(* IEC 61131-3 sources: Codesys_IAP/Demo/PLC1/Magazijn Overzetter Simulatie Structured Text 2V1_tekst/Programma Structured Text/StationClass, 8 files *)

(* ---- cycle.st ---- *)
(*#### DECLARATIE ####*)
// Datum : 26 november 2026, Auteur: Gerard Harkema
METHOD cycle
VAR
END_VAR
(*#### IMPLEMENTATIE ####*)
// Eerst de objecten
magazijn.cycle();
overzetter.cycle();

// Dan de fouten: een fout in een object zet het hele station in error
IF magazijn.isError() OR overzetter.isError() THEN
	eState := stationStates.error;
END_IF

// Dan de coordinatie, volgens het statediagram van StationClass
CASE eState OF
	stationStates.idle:
		; // wacht op start()

	stationStates.magazijn_uitstoten:
		IF magazijn.start() THEN		// TRUE = mislukt
			eState := stationStates.error;
		ELSE
			eState := stationStates.wacht_magazijn_klaar;
		END_IF

	stationStates.wacht_magazijn_klaar:
		IF magazijn.isKlaar() THEN
			eState := stationStates.overzetten;
		END_IF

	stationStates.overzetten:
		IF overzetter.start() THEN		// TRUE = mislukt
			eState := stationStates.error;
		ELSE
			eState := stationStates.wacht_overzetter_klaar;
		END_IF

	stationStates.wacht_overzetter_klaar:
		IF overzetter.isKlaar() THEN
			eState := stationStates.idle;
		END_IF

	stationStates.error:
		; // wacht op reset()
END_CASE

(* ---- initialize.st ---- *)
(*#### DECLARATIE ####*)
// Datum : 26 november 2026, Auteur: Gerard Harkema
METHOD initialize
VAR_INPUT
	IORef			: REFERENCE TO stationIO;
END_VAR
(*#### IMPLEMENTATIE ####*)
IO REF= IORef;

// Elk object krijgt zijn eigen IO-structuur
magazijn.initialize(IO.magazijn);
overzetter.initialize(IO.overzetter);

eState := stationStates.idle;

(* ---- isError.st ---- *)
(*#### DECLARATIE ####*)
// Datum : 26 november 2026, Auteur: Gerard Harkema
METHOD isError : BOOL
VAR_INPUT
END_VAR
(*#### IMPLEMENTATIE ####*)
isError := (eState = stationStates.error);

(* ---- isKlaar.st ---- *)
(*#### DECLARATIE ####*)
// Datum : 26 november 2026, Auteur: Gerard Harkema
METHOD isKlaar : BOOL
VAR_INPUT
END_VAR
(*#### IMPLEMENTATIE ####*)
isKlaar := (eState = stationStates.idle)
		AND magazijn.isKlaar()
		AND overzetter.isKlaar();

(* ---- isMagazijnLeeg.st ---- *)
(*#### DECLARATIE ####*)
// Datum : 26 november 2026, Auteur: Gerard Harkema
METHOD isMagazijnLeeg : BOOL
VAR_INPUT
END_VAR
(*#### IMPLEMENTATIE ####*)
isMagazijnLeeg := magazijn.isMagazijnLeeg();

(* ---- noodstop.st ---- *)
(*#### DECLARATIE ####*)
// Datum : 26 november 2026, Auteur: Gerard Harkema
METHOD noodstop
VAR_INPUT
END_VAR
(*#### IMPLEMENTATIE ####*)
// Noodstop geeft het station door aan beide objecten
magazijn.noodstop();
overzetter.noodstop();
eState := stationStates.error;

(* ---- reset.st ---- *)
(*#### DECLARATIE ####*)
// Datum : 26 november 2026, Auteur: Gerard Harkema
METHOD reset
VAR_INPUT
END_VAR
(*#### IMPLEMENTATIE ####*)
// Reset geeft het station door aan beide objecten; die gaan eerst naar hun veilige stand
magazijn.reset();
overzetter.reset();
eState := stationStates.idle;

(* ---- start.st ---- *)
(*#### DECLARATIE ####*)
// Datum : 26 november 2026, Auteur: Gerard Harkema
METHOD start : BOOL
VAR_INPUT
END_VAR
(*#### IMPLEMENTATIE ####*)
// Start een cyclus: een beker uit het magazijn naar de afgifteplaats.
// Kan alleen vanuit idle en als beide objecten in hun ruststand staan.
IF NOT isKlaar() THEN
	start := TRUE; // Failed (station blijft gewoon doorgaan met wat het deed)
	RETURN;
END_IF

eState := stationStates.magazijn_uitstoten;
start := FALSE; // oké
